(* PLC project Vn_ld_neg_contact, Beckhoff Automation GmbH TwinCAT PLC Control 3.5.13.21 *)
(* stored: creationDateTime 1970-01-01T00:00:00 *)

PROGRAM Vn_ld_neg_contact

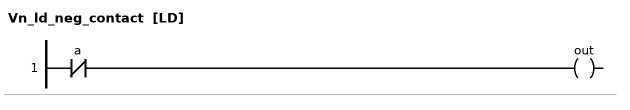
(* LD diagram, written out as Structured Text *)
out := NOT a;
END_PROGRAM
